// TIA Portal V20 export
// export: Created 2026-10-12T16:46:21.4659687Z, ExportSetting WithDefaults, DisplayName Totally Integrated Automation Portal, DisplayVersion V20 Update 6, DisplayName TIA Portal Openness, DisplayVersion V20 Update 6, DisplayName TIA Portal Version Control Interface, DisplayVersion V20 Update 6, DisplayName SINAMICS Startdrive Advanced, DisplayVersion V20 SP1 Update 2, DisplayName SINAMICS Startdrive G110M, G120, G120C, G120D, G120P, G115D, DisplayVersion V20 SP1 Update 2, DisplayName SINAMICS Startdrive G130, G150, S120, S150, SINAMICS MV, G220, S200, S210, DisplayVersion V20 SP1 Update 2, DisplayName STEP 7 Professional, DisplayVersion V20 Update 6, DisplayName STEP 7 Safety, DisplayVersion V20 Update 2, DisplayName WinCC Basic/Comfort/Advanced, DisplayVersion V20 Update 6, DisplayName WinCC Professional, DisplayVersion V20 Update 6, DisplayName WinCC Unified, DisplayVersion V20 Update 6
DATA_BLOCK "FB_FlexKraft_DB"   // DB6
VERSION : 0.1
// stored: AutoNumber true, DBAccessibleFromOPCUA true, DBAccessibleFromWebserver true, InstanceOfName FB_FlexKraft, InstanceOfType FB
"FB_FlexKraft"
   // VAR_INPUT
   //    bOn : Bool;
   //    bStartA : Bool;
   //    bBlockA : Bool;
   //    bRunProgA : Bool;
   //    bReverseA : Bool;
   //    bReverseB : Bool;
   //    bStartB : Bool;
   //    bClrAhA : Bool;
   //    bClrAhB : Bool;
   //    bClrTimer : Bool;
   //    bBlockB : Bool;
   //    bAuxOutA : Bool;
   //    bAuxOutB : Bool;
   //    bRunProgB : Bool;
   //    iSetVoltage_cV : Int;
   //    iSetCurrent_raw : Int;
   //    wStartramp_dS : Word;
   // END_VAR
   // VAR_OUTPUT
   //    bAlarm : Bool;
   //    bWarning : Bool;
   //    bRemote : Bool;
   //    bRunningA : Bool;
   //    bAhLimitA : Bool;
   //    bAhLimitB : Bool;
   //    bTimerLimitA : Bool;
   //    bVoltageModeA : Bool;
   //    bVoltageModeB : Bool;
   //    bUnitOn : Bool;
   //    bHiRes : Bool;
   //    bRunningB : Bool;
   //    iOutVoltage_cV : Int;
   //    iOutCurrent_raw : Int;
   //    wWarnings : Word;
   //    wAlarms : Word;
   // END_VAR
   // VAR_IN_OUT
   //    stDev : "UDT_FlexKraft_Device";
   // END_VAR
BEGIN
END_DATA_BLOCK
